SUBAPPLICATION Uebung_163 (* Übung zu logiBUS_ENC_ID und logiBUS_QW_SERVO: Servo mit dem Drehgeber stellen *)
  (* Standard: 61499-2; Description: Copyright (c) 2026 Meisterschulen am Ostbahnhof This program and the accompanying materials are made available under the terms of the Eclipse Public License 2.0 which is available at https://www.eclipse.org/legal/epl-2.0/ SPDX-License-Identifier: EPL-2.0 *)
  (* Version 1.0, 2026-11-26, Franz Höpfinger, Meisterschulen am Ostbahnhof, initial API and implementation and/or initial documentation *)
  PACKAGE Uebungen;
  IMPORT Uebungen::const::UT::DefaultPool::OutputNumber_N1;
  IMPORT logiBUS::io::ENC::logiBUS_ENC::Encoder_E1;
  IMPORT logiBUS::io::DI::logiBUS_DI::Input_I9;
  IMPORT logiBUS::io::DI::logiBUS_DI_Events::BUTTON_SINGLE_CLICK;
  IMPORT logiBUS::io::DQ::logiBUS_DO::Output_Q1;
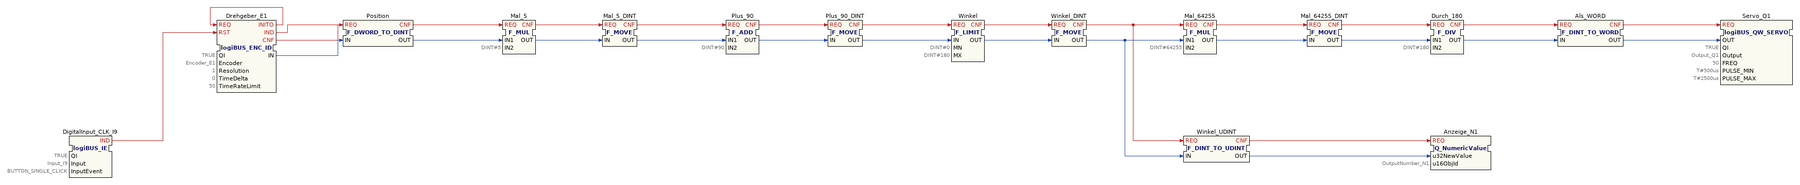
  (* Servo mit dem Inkrementalgeber stellen (Trainer20: Drehgeber A = GPIO22, B = GPIO23, Taster = I9, Servo an Q1). Position 0 = Mitte 90 Grad. Je Raste 5 Grad: ins Minus Richtung 0 Grad, ins Plus Richtung 180 Grad. F_LIMIT hält den Winkel zwischen 0 und 180 Grad. Winkel * 64255 / 180 ergibt OUT (0..16#FAFF) für logiBUS_QW_SERVO. Der Winkel steht am VT auf OutputNumber N1. Beim Start fragt INITO die Position einmal ab, der Servo fährt auf 90 Grad. I9 Klick: RST, zurück auf 90 Grad. PULSE_MIN/PULSE_MAX (hier 500/2500 us für 0/180 Grad) laut Datenblatt des Servos anpassen. Viele Servos machen mit 1000/2000 us nur etwa 90 Grad Weg. *)
  FBS
    Drehgeber_E1 : logiBUS::io::ENC::logiBUS_ENC_ID(QI := TRUE, Encoder := Encoder_E1, Resolution := 1, TimeDelta := 0, TimeRateLimit := 50); (* Trainer20: A = GPIO22, B = GPIO23 *)
    Position : iec61131::conversion::F_DWORD_TO_DINT;
    Mal_5 : iec61131::arithmetic::F_MUL(IN2 := DINT#5); (* 5 Grad je Raste *)
    Mal_5_DINT : iec61131::selection::F_MOVE; {SET_ATTRIBUTE(DataType, DINT)}
    Plus_90 : iec61131::arithmetic::F_ADD(IN2 := DINT#90); (* Position 0 = Mitte 90 Grad *)
    Plus_90_DINT : iec61131::selection::F_MOVE; {SET_ATTRIBUTE(DataType, DINT)}
    Winkel : iec61131::selection::F_LIMIT(MN := DINT#0, MX := DINT#180); (* 0 bis 180 Grad *)
    Winkel_DINT : iec61131::selection::F_MOVE; {SET_ATTRIBUTE(DataType, DINT)}
    Mal_64255 : iec61131::arithmetic::F_MUL(IN2 := DINT#64255); (* 180 Grad = 16#FAFF *)
    Mal_64255_DINT : iec61131::selection::F_MOVE; {SET_ATTRIBUTE(DataType, DINT)}
    Durch_180 : iec61131::arithmetic::F_DIV(IN2 := DINT#180);
    Als_WORD : iec61131::conversion::F_DINT_TO_WORD;
    Servo_Q1 : logiBUS::io::DO_SERVO::logiBUS_QW_SERVO(QI := TRUE, Output := Output_Q1, FREQ := 50, PULSE_MIN := T#500us, PULSE_MAX := T#2500us); (* 0 Grad = PULSE_MIN, 180 Grad = PULSE_MAX *)
    Winkel_UDINT : iec61131::conversion::F_DINT_TO_UDINT;
    Anzeige_N1 : isobus::UT::Q::Q_NumericValue(u16ObjId := OutputNumber_N1); (* Winkel in Grad am VT *)
    DigitalInput_CLK_I9 : logiBUS::io::DI::logiBUS_IE(QI := TRUE, Input := Input_I9, InputEvent := BUTTON_SINGLE_CLICK); (* Taster am Drehgeber: zurück auf 90 Grad *)
  END_FBS
  EVENT_CONNECTIONS
    Drehgeber_E1.INITO TO Drehgeber_E1.REQ;
    Drehgeber_E1.IND TO Position.REQ;
    Drehgeber_E1.CNF TO Position.REQ;
    Position.CNF TO Mal_5.REQ;
    Mal_5_DINT.CNF TO Plus_90.REQ;
    Plus_90_DINT.CNF TO Winkel.REQ;
    Winkel_DINT.CNF TO Mal_64255.REQ;
    Mal_64255_DINT.CNF TO Durch_180.REQ;
    Durch_180.CNF TO Als_WORD.REQ;
    Als_WORD.CNF TO Servo_Q1.REQ;
    Winkel_DINT.CNF TO Winkel_UDINT.REQ;
    Winkel_UDINT.CNF TO Anzeige_N1.REQ;
    DigitalInput_CLK_I9.IND TO Drehgeber_E1.RST;
    Mal_5.CNF TO Mal_5_DINT.REQ;
    Plus_90.CNF TO Plus_90_DINT.REQ;
    Winkel.CNF TO Winkel_DINT.REQ;
    Mal_64255.CNF TO Mal_64255_DINT.REQ;
  END_CONNECTIONS
  DATA_CONNECTIONS
    Drehgeber_E1.IN TO Position.IN;
    Position.OUT TO Mal_5.IN1;
    Mal_5_DINT.OUT TO Plus_90.IN1;
    Plus_90_DINT.OUT TO Winkel.IN;
    Winkel_DINT.OUT TO Mal_64255.IN1;
    Mal_64255_DINT.OUT TO Durch_180.IN1;
    Durch_180.OUT TO Als_WORD.IN;
    Als_WORD.OUT TO Servo_Q1.OUT;
    Winkel_DINT.OUT TO Winkel_UDINT.IN;
    Winkel_UDINT.OUT TO Anzeige_N1.u32NewValue;
    Mal_5.OUT TO Mal_5_DINT.IN;
    Plus_90.OUT TO Plus_90_DINT.IN;
    Winkel.OUT TO Winkel_DINT.IN;
    Mal_64255.OUT TO Mal_64255_DINT.IN;
  END_CONNECTIONS
END_SUBAPPLICATION
